// TwinCAT 3 PLC project TestSample
// ProgramVersion: 3.1.4026.28
// libraries:
//   Tc2_Standard, * (Beckhoff Automation GmbH)
//   Tc2_System, * (Beckhoff Automation GmbH)
//   Tc2_TcpIp, * (Beckhoff Automation GmbH)
//   Tc3_Module, * (Beckhoff Automation GmbH)
// project tree:
//   Diagram/ Class Diagram.TcCD (not stored)
//   Generated/DUT_Generated/ ST_VC_InspectionResult.TcDUT, ST_VC_MoveToPositionArgs.TcDUT, ST_VC_MoveToPositionResult.TcDUT, ST_VC_ReportModuleStateArgs.TcDUT
//   Generated/GVLs_Generated/ GVL_VC_Methods.TcGVL
//   Generated/POU_Generated/ VC_Call_StartInspection.TcPOU, VC_Handle_MoveToPosition.TcPOU, VC_Handle_ReportModuleState.TcPOU
//   Library/DUT/ E_VC_LinkState.TcDUT, E_VC_MsgType.TcDUT, E_VC_SlotState.TcDUT, ST_VC_CtrlMsg.TcDUT, ST_VC_Diag.TcDUT, ST_VC_Header.TcDUT, ST_VC_InSlot.TcDUT, ST_VC_LinkData.TcDUT, ST_VC_MethodInfo.TcDUT, ST_VC_OutSlot.TcDUT
//   Library/GVL/ GVL_VC_Param.TcGVL
//   Library/POU/ VC_CancelOutSlot.TcPOU, VC_CompleteInSlot.TcPOU, VC_DecodeHeader.TcPOU, VC_EncodeHeader.TcPOU, VC_Framer.TcPOU, VC_GetBool.TcPOU, VC_GetFloat32.TcPOU, VC_GetFloat32Array.TcPOU, VC_GetFloat64.TcPOU, VC_GetInt16.TcPOU, VC_GetInt32.TcPOU, VC_GetInt64.TcPOU, VC_GetInt8.TcPOU, VC_GetRaw.TcPOU, VC_GetString.TcPOU, VC_GetUInt16.TcPOU, VC_GetUInt32.TcPOU, VC_GetUInt64.TcPOU, VC_GetUInt8.TcPOU, VC_IsCallable.TcPOU, VC_Link.TcPOU, VC_MethodIndex.TcPOU, VC_PutBool.TcPOU, VC_PutFloat32.TcPOU, VC_PutFloat32Array.TcPOU, VC_PutFloat64.TcPOU, VC_PutInt16.TcPOU, VC_PutInt32.TcPOU, VC_PutInt64.TcPOU, VC_PutInt8.TcPOU, VC_PutRaw.TcPOU, VC_PutString.TcPOU, VC_PutUInt16.TcPOU, VC_PutUInt32.TcPOU, VC_PutUInt64.TcPOU, VC_PutUInt8.TcPOU, VC_ReleaseOutSlot.TcPOU, VC_ReserveOutSlot.TcPOU, VC_SubmitOutSlot.TcPOU, VC_TakeInSlot.TcPOU, VC_Transport.TcPOU
//   / PlcTask.TcTTO
//   POUs/ MAIN.TcPOU
//   Test/GVL/ GVL_VC.TcGVL
//   Test/POU/ FB_VC_LinkTest.TcPOU, MAIN_1.TcPOU
// real-time tasks:
//   TASK PlcTask: cycle T#10ms, priority 20, ADS port 350

CONFIGURATION TestSample
    RESOURCE PLC ON TwinCAT3
        TASK PlcTask(INTERVAL := T#10ms, PRIORITY := 20);
    END_RESOURCE
END_CONFIGURATION

// ---- Generated/DUT_Generated/ST_VC_InspectionResult.TcDUT
TYPE ST_VC_InspectionResult :
STRUCT
    Pass          : BOOL;
    ErrorCode     : DINT;
    MeasuredCount : UINT;
    Measured      : ARRAY[0..15] OF REAL;
END_STRUCT
END_TYPE

// ---- Generated/DUT_Generated/ST_VC_MoveToPositionArgs.TcDUT
TYPE ST_VC_MoveToPositionArgs :
STRUCT
    Position : LREAL;
END_STRUCT
END_TYPE

// ---- Generated/DUT_Generated/ST_VC_MoveToPositionResult.TcDUT
TYPE ST_VC_MoveToPositionResult :
STRUCT
    Accepted : BOOL;
END_STRUCT
END_TYPE

// ---- Generated/DUT_Generated/ST_VC_ReportModuleStateArgs.TcDUT
TYPE ST_VC_ReportModuleStateArgs :
STRUCT
    State   : UINT;     // PackML state from VisionCore
    AlarmId : DINT;
END_STRUCT
END_TYPE

// ---- Library/DUT/E_VC_LinkState.TcDUT
TYPE E_VC_LinkState :
(
    VC_LS_DISABLED   := 0,
    VC_LS_CONNECTING := 1,   // PLC connects actively (VisionCore mode Listen)
    VC_LS_LISTENING  := 2,   // PLC waits for connection (VisionCore mode Connect)
    VC_LS_HELLO      := 3,   // Hello sent, waiting for HelloAck
    VC_LS_ONLINE     := 4,
    VC_LS_CLOSING    := 5,
    VC_LS_WAIT_RETRY := 6
) UINT;
END_TYPE

// ---- Library/DUT/E_VC_MsgType.TcDUT
TYPE E_VC_MsgType :
// Deliberately NOT {attribute 'strict'}: values are compared with the USINT header field.
(
    VC_MT_HELLO     := 1,
    VC_MT_HELLO_ACK := 2,
    VC_MT_REQUEST   := 3,
    VC_MT_RESPONSE  := 4,
    VC_MT_CANCEL    := 5,
    VC_MT_HEARTBEAT := 6
) USINT;
END_TYPE

// ---- Library/DUT/E_VC_SlotState.TcDUT
TYPE E_VC_SlotState :
(
    VC_SS_FREE           := 0,
    VC_SS_RESERVED       := 1,   // Out: block owns slot
    VC_SS_TX_PENDING     := 2,   // Out: request ready to send
    VC_SS_SENT           := 3,   // Out: request sent, waiting for response
    VC_SS_CANCEL_PENDING := 4,   // Out: Cancel must be sent
    VC_SS_DONE           := 5,   // Out: response or error available
    VC_SS_REQUEST        := 10,  // In:  request received, no handler yet
    VC_SS_IN_PROGRESS    := 11,  // In:  handler working
    VC_SS_RESPONSE_READY := 12   // In:  response ready to send
) UINT;
END_TYPE

// ---- Library/DUT/ST_VC_CtrlMsg.TcDUT
TYPE ST_VC_CtrlMsg :              // Cancel or error response without payload
STRUCT
    MessageType : E_VC_MsgType;
    MethodId    : UINT;
    CallId      : UDINT;
    Status      : UINT;
END_STRUCT
END_TYPE

// ---- Library/DUT/ST_VC_Diag.TcDUT
TYPE ST_VC_Diag :
STRUCT
    RxMessages          : UDINT;
    TxMessages          : UDINT;
    ProtocolErrors      : UDINT;
    Reconnects          : UDINT;
    CallTimeouts        : UDINT;
    RejectedCalls       : UDINT;
    LastErrorId         : UINT;
    LastErrorMs         : UDINT;
    LastTransportStatus : DWORD;  // raw nErrId of the Tc2_TcpIp block
END_STRUCT
END_TYPE

// ---- Library/DUT/ST_VC_Header.TcDUT
{attribute 'pack_mode' := '1'}
TYPE ST_VC_Header :
STRUCT
    Magic           : UINT;    // 16#5643, little-endian on the wire (43 56)
    ProtocolVersion : USINT;   // 1
    MessageType     : USINT;   // E_VC_MsgType
    Flags           : UINT;    // reserved, 0
    MethodId        : UINT;    // 0 for Hello / Heartbeat
    CallId          : UDINT;   // bit 31 = 1: call from VisionCore
    PayloadLength   : UDINT;
    Status          : UINT;    // response status, else 0
    Reserved        : UINT;
END_STRUCT
END_TYPE

// ---- Library/DUT/ST_VC_InSlot.TcDUT
TYPE ST_VC_InSlot :               // App calls PLC
STRUCT
    State           : E_VC_SlotState;
    MethodIndex     : UINT;
    CallId          : UDINT;
    ReceivedMs      : UDINT;
    CancelRequested : BOOL;
    Status          : UINT;
    PayloadLen      : UDINT;
    Payload         : ARRAY[0..VC_MAX_PAYLOAD - 1] OF BYTE;  // arguments first, then result
END_STRUCT
END_TYPE

// ---- Library/DUT/ST_VC_LinkData.TcDUT
TYPE ST_VC_LinkData :
STRUCT
    // State
    State          : E_VC_LinkState;
    Online         : BOOL;
    NowMs          : UDINT;      // time base, set by VC_Link every cycle
    StateSinceMs   : UDINT;
    LastRxMs       : UDINT;
    LastTxMs       : UDINT;
    NextCallId     : UDINT;      // 1 .. 16#7FFFFFFF, bit 31 always 0

    // Release from HelloAck and handler presence, index = method index
    MethodState    : ARRAY[0..VC_MAX_METHODS - 1] OF USINT;  // 0 unknown, 1 released, 2 hash, 3 not allowed
    HandlerSeenMs  : ARRAY[0..VC_MAX_METHODS - 1] OF UDINT;

    // Call slots
    OutSlots       : ARRAY[0..VC_MAX_CALLS - 1] OF ST_VC_OutSlot;
    InSlots        : ARRAY[0..VC_MAX_CALLS - 1] OF ST_VC_InSlot;
    NextOutSend    : UINT;       // round robin for sending

    // Control messages
    CtrlQueue      : ARRAY[0..VC_CTRL_QUEUE - 1] OF ST_VC_CtrlMsg;
    CtrlHead       : UINT;
    CtrlCount      : UINT;

    // Buffers
    RxBuffer       : ARRAY[0..VC_RX_BUFFER - 1] OF BYTE;
    RxFill         : UDINT;
    TxFrame        : ARRAY[0..VC_HEADER_LEN + VC_MAX_PAYLOAD - 1] OF BYTE;

    // Diagnostics
    Diag           : ST_VC_Diag;
END_STRUCT
END_TYPE

// ---- Library/DUT/ST_VC_MethodInfo.TcDUT
TYPE ST_VC_MethodInfo :
STRUCT
    MethodId  : UINT;
    Hash      : UDINT;   // CRC-32 of canonical signature (generated)
    Provider  : USINT;   // 0 = App, 1 = Plc
    TimeoutMs : UDINT;
    ArgsLen   : UDINT;   // request payload length
    ResultLen : UDINT;   // response payload length at status 0
END_STRUCT
END_TYPE

// ---- Library/DUT/ST_VC_OutSlot.TcDUT
TYPE ST_VC_OutSlot :              // PLC calls App
STRUCT
    State        : E_VC_SlotState;
    MethodIndex  : UINT;
    CallId       : UDINT;
    StartMs      : UDINT;
    TimeoutMs    : UDINT;
    OwnerSeenMs  : UDINT;         // last call of owning VC_Call_* block
    Status       : UINT;
    PayloadLen   : UDINT;
    Payload      : ARRAY[0..VC_MAX_PAYLOAD - 1] OF BYTE;  // arguments first, then result
END_STRUCT
END_TYPE

// ---- Generated/GVLs_Generated/GVL_VC_Methods.TcGVL
VAR_GLOBAL CONSTANT
// ===== GENERATED PART (normally written by vcgen) - hand-written stand-in for testing =====
// Hash = CRC-32 (IEEE, as zlib) over the canonical signature, SPS-Konzept 4.5:
//   10|StartInspection|App|UInt16,String32|Bool,Int32,UInt16,Float32[16]
//   500|ReportModuleState|Plc|UInt16,Int32|
//   600|MoveToPosition|Plc|Float64|Bool
// ASSUMPTION: VisionCore computes the same CRC variant and string. If not, HelloAck returns
// MethodState 2 and calls fail with ErrorId 2 -> copy the hashes from the VisionCore build.
    VC_METHOD_COUNT            : UINT := 3;

    // Method index = position in VC_METHODS (used by all blocks)
    VC_IDX_START_INSPECTION    : UINT := 0;
    VC_IDX_REPORT_MODULE_STATE : UINT := 1;
    VC_IDX_MOVE_TO_POSITION    : UINT := 2;

    // ASSUMPTION: project interface name, confirm with VisionCore configuration
    VC_INTERFACES : ARRAY[0..3] OF STRING(47) := ['VisionCore.Platform', 'Stent.Line1', '', ''];

    VC_METHODS : ARRAY[0..VC_MAX_METHODS - 1] OF ST_VC_MethodInfo := [
        // StartInspection: args UInt16 + String32 = 34; result Bool+Int32+UInt16+16xFloat32 = 71
        (MethodId := 10,  Hash := 16#A1EFD4EB, Provider := 0, TimeoutMs := 10000, ArgsLen := 34, ResultLen := 71),
        // ReportModuleState: args UInt16 + Int32 = 6; no result
        (MethodId := 500, Hash := 16#18245D80, Provider := 1, TimeoutMs := 200,   ArgsLen := 6,  ResultLen := 0),
        // MoveToPosition: args Float64 = 8; result Bool = 1. ASSUMPTION: timeout 5000 ms
        (MethodId := 600, Hash := 16#689DF4EB, Provider := 1, TimeoutMs := 5000,  ArgsLen := 8,  ResultLen := 1)
    ];
END_VAR

// ---- Library/GVL/GVL_VC_Param.TcGVL
VAR_GLOBAL CONSTANT
    // ---- Protocol (fixed, SPS-Konzept section 5) ----
    VC_MAGIC              : UINT  := 16#5643;   // 'VC'
    VC_PROTOCOL_VERSION   : USINT := 1;
    VC_HEADER_LEN         : UDINT := 20;
    VC_HELLO_ACK_LEN      : UDINT := 65;        // Accepted + 64 x MethodState
    VC_PROVIDER_APP       : USINT := 0;
    VC_PROVIDER_PLC       : USINT := 1;

    // ---- Parameters (Bausteindesign section 3) ----
    VC_MAX_PAYLOAD        : UDINT := 4096;
    VC_MAX_CALLS          : UINT  := 8;
    VC_MAX_METHODS        : UINT  := 64;        // must stay 64: Hello/HelloAck carry 64 entries
    VC_RX_BUFFER          : UDINT := 2 * (VC_HEADER_LEN + VC_MAX_PAYLOAD);
    VC_CTRL_QUEUE         : UINT  := 16;
    VC_MSG_PER_CYCLE      : UINT  := 4;
    VC_HELLO_TIMEOUT_MS   : UDINT := 5000;
    VC_HEARTBEAT_MS       : UDINT := 1000;
    VC_WATCHDOG_MS        : UDINT := 3000;
    VC_RETRY_MS           : UDINT := 2000;
    VC_OWNER_TIMEOUT_MS   : UDINT := 1000;

    // ---- Status codes (SPS-Konzept 5.7) ----
    VC_STATUS_OK                  : UINT := 0;
    VC_STATUS_UNKNOWN_METHOD      : UINT := 1;
    VC_STATUS_METHOD_INCOMPATIBLE : UINT := 2;
    VC_STATUS_NOT_ALLOWED         : UINT := 3;
    VC_STATUS_INVALID_PAYLOAD     : UINT := 4;
    VC_STATUS_BUSY                : UINT := 5;
    VC_STATUS_CANCELLED           : UINT := 6;
    VC_STATUS_TIMEOUT             : UINT := 7;
    VC_STATUS_CONNECTION_LOST     : UINT := 8;
    VC_STATUS_INTERNAL_ERROR      : UINT := 9;

    // ---- VC_Link.ErrorId (Bausteindesign section 8) ----
    VC_ERR_CONNECT         : UINT := 1;   // connect / listen / accept failed
    VC_ERR_HELLO_TIMEOUT   : UINT := 2;   // no HelloAck in time
    VC_ERR_HELLO_REJECTED  : UINT := 3;   // HelloAck Accepted = FALSE
    VC_ERR_PROTOCOL        : UINT := 4;   // invalid header / unexpected message
    VC_ERR_WATCHDOG        : UINT := 5;   // nothing received
    VC_ERR_SEND            : UINT := 6;
    VC_ERR_RECEIVE         : UINT := 7;
END_VAR

// ---- Test/GVL/GVL_VC.TcGVL
VAR_GLOBAL
    LinkData : ST_VC_LinkData;   // one per VisionCore connection, ~80 KB
END_VAR

// ---- Library/POU/VC_Link.TcPOU
FUNCTION_BLOCK VC_Link
// Central block: one instance per VisionCore connection, called every cycle,
// BEFORE all VC_Call_* / VC_Handle_* blocks that use the same ST_VC_LinkData (same task).
VAR_INPUT
    Enable        : BOOL;
    Mode          : INT;           // 0 = connect actively, 1 = wait for connection
    RemoteAddress : STRING(15);    // Mode = 0
    RemotePort    : UINT := 5100;  // Mode = 0
    LocalPort     : UINT := 5100;  // Mode = 1
    ClientId      : STRING(31);
END_VAR
VAR_IN_OUT
    Link          : ST_VC_LinkData;
END_VAR
VAR_OUTPUT
    Connected     : BOOL;          // TCP connection up
    Online        : BOOL;          // HelloAck received
    Restricted    : BOOL;          // at least one method not released
    Error         : BOOL;          // stays set until ONLINE again
    ErrorId       : UINT;          // VC_ERR_*
    State         : E_VC_LinkState;
END_VAR
VAR
    fbTransport   : VC_Transport;
    fbFramer      : VC_Framer;
    bSendReq      : BOOL;          // frame in TxFrame, waiting for transport to take it
    nTxLen        : UDINT;
    bHelloSent    : BOOL;
    nIdx          : UINT;
END_VAR

// ---- 1. Time base ----
Link.NowMs := TIME_TO_UDINT(TIME());

// ---- 2./3. Transport: connect, accept, close, send, receive ----
fbTransport(
    Open          := (Link.State = VC_LS_CONNECTING) OR (Link.State = VC_LS_LISTENING)
                     OR (Link.State = VC_LS_HELLO) OR (Link.State = VC_LS_ONLINE),
    Mode          := Mode,
    RemoteAddress := RemoteAddress,
    RemotePort    := RemotePort,
    LocalPort     := LocalPort,
    SendRequest   := bSendReq,
    SendLen       := nTxLen,
    Link          := Link);
IF fbTransport.SendBusy THEN
    bSendReq := FALSE;                 // transport has taken the frame
END_IF
IF fbTransport.Error THEN
    Link.Diag.LastTransportStatus := fbTransport.Status;
END_IF

// ---- Connection state machine ----
CASE Link.State OF
VC_LS_DISABLED:
    IF Enable THEN
        IF Mode = 0 THEN
            THIS^.GotoState(stLink := Link, NewState := VC_LS_CONNECTING);
        ELSE
            THIS^.GotoState(stLink := Link, NewState := VC_LS_LISTENING);
        END_IF
    END_IF

VC_LS_CONNECTING, VC_LS_LISTENING:
    IF NOT Enable THEN
        THIS^.GotoState(stLink := Link, NewState := VC_LS_CLOSING);
    ELSIF fbTransport.Error THEN
        THIS^.SetError(stLink := Link, Id := VC_ERR_CONNECT);
        THIS^.GotoState(stLink := Link, NewState := VC_LS_CLOSING);   // releases handles, then WAIT_RETRY
    ELSIF fbTransport.Connected THEN
        THIS^.GotoState(stLink := Link, NewState := VC_LS_HELLO);
    END_IF

VC_LS_HELLO, VC_LS_ONLINE:
    IF NOT Enable THEN
        THIS^.GotoState(stLink := Link, NewState := VC_LS_CLOSING);
    ELSIF fbTransport.Error THEN
        THIS^.SetError(stLink := Link, Id := fbTransport.ErrorId);
        THIS^.GotoState(stLink := Link, NewState := VC_LS_CLOSING);
    ELSIF NOT fbTransport.Connected THEN
        THIS^.SetError(stLink := Link, Id := VC_ERR_RECEIVE);
        THIS^.GotoState(stLink := Link, NewState := VC_LS_CLOSING);
    END_IF

VC_LS_CLOSING:
    IF fbTransport.Idle THEN
        IF Enable THEN
            THIS^.GotoState(stLink := Link, NewState := VC_LS_WAIT_RETRY);
        ELSE
            THIS^.GotoState(stLink := Link, NewState := VC_LS_DISABLED);
        END_IF
    END_IF

VC_LS_WAIT_RETRY:
    IF NOT Enable THEN
        THIS^.GotoState(stLink := Link, NewState := VC_LS_DISABLED);
    ELSIF (Link.NowMs - Link.StateSinceMs) >= VC_RETRY_MS THEN
        IF Mode = 0 THEN
            THIS^.GotoState(stLink := Link, NewState := VC_LS_CONNECTING);
        ELSE
            THIS^.GotoState(stLink := Link, NewState := VC_LS_LISTENING);
        END_IF
    END_IF
END_CASE

// ---- 4. Process messages ----
IF (Link.State = VC_LS_HELLO) OR (Link.State = VC_LS_ONLINE) THEN
    THIS^.ProcessMessages(stLink := Link);
END_IF

// ---- 5. Deadlines ----
IF (Link.State = VC_LS_HELLO) OR (Link.State = VC_LS_ONLINE) THEN
    THIS^.CheckDeadlines(stLink := Link);
END_IF

// ---- 6. Schedule at most one message ----
IF (Link.State = VC_LS_HELLO) OR (Link.State = VC_LS_ONLINE) THEN
    THIS^.ScheduleSend(stLink := Link);
END_IF

// ---- 7. Outputs ----
Connected  := fbTransport.Connected;
Online     := Link.Online;
State      := Link.State;
Restricted := FALSE;
IF Link.Online THEN
    nIdx := 0;
    WHILE (nIdx < VC_METHOD_COUNT) AND (nIdx < VC_MAX_METHODS) DO
        IF Link.MethodState[nIdx] <> 1 THEN
            Restricted := TRUE;
        END_IF
        nIdx := nIdx + 1;
    END_WHILE
END_IF

METHOD PRIVATE BuildHello : UDINT
// Bausteindesign 7.3: 32 + 4 x 48 + 2 + 64 x 6 = 610 bytes payload
VAR_IN_OUT
    stLink : ST_VC_LinkData;
END_VAR
VAR
    nPos : UDINT;
    k    : UINT;
END_VAR
nPos := VC_HEADER_LEN;
VC_PutString(Buf := stLink.TxFrame, Pos := nPos, Value := ClientId, Len := 32);
FOR k := 0 TO 3 DO
    VC_PutString(Buf := stLink.TxFrame, Pos := nPos, Value := VC_INTERFACES[k], Len := 48);
END_FOR
VC_PutUInt16(Buf := stLink.TxFrame, Pos := nPos, Value := VC_METHOD_COUNT);
FOR k := 0 TO VC_MAX_METHODS - 1 DO
    VC_PutUInt16(Buf := stLink.TxFrame, Pos := nPos, Value := VC_METHODS[k].MethodId);
    VC_PutUInt32(Buf := stLink.TxFrame, Pos := nPos, Value := VC_METHODS[k].Hash);
END_FOR
BuildHello := nPos - VC_HEADER_LEN;
END_METHOD

METHOD PRIVATE CheckDeadlines
VAR_IN_OUT
    stLink : ST_VC_LinkData;
END_VAR
VAR
    k    : UINT;
    nIdx : UINT;
END_VAR
// Hello timeout / watchdog
IF stLink.State = VC_LS_HELLO THEN
    IF (stLink.NowMs - stLink.StateSinceMs) > VC_HELLO_TIMEOUT_MS THEN
        THIS^.SetError(stLink := stLink, Id := VC_ERR_HELLO_TIMEOUT);
        THIS^.GotoState(stLink := stLink, NewState := VC_LS_CLOSING);
        RETURN;
    END_IF
ELSIF stLink.State = VC_LS_ONLINE THEN
    IF (stLink.NowMs - stLink.LastRxMs) > VC_WATCHDOG_MS THEN
        THIS^.SetError(stLink := stLink, Id := VC_ERR_WATCHDOG);
        THIS^.GotoState(stLink := stLink, NewState := VC_LS_CLOSING);
        RETURN;
    END_IF
END_IF

FOR k := 0 TO VC_MAX_CALLS - 1 DO
    // Out slots: call timeout and orphaned slots
    CASE stLink.OutSlots[k].State OF
    VC_SS_SENT:
        IF (stLink.NowMs - stLink.OutSlots[k].StartMs) > stLink.OutSlots[k].TimeoutMs THEN
            stLink.OutSlots[k].Status := VC_STATUS_TIMEOUT;
            stLink.OutSlots[k].State  := VC_SS_CANCEL_PENDING;
            stLink.Diag.CallTimeouts  := stLink.Diag.CallTimeouts + 1;
        END_IF
    VC_SS_RESERVED, VC_SS_DONE:
        IF (stLink.NowMs - stLink.OutSlots[k].OwnerSeenMs) > VC_OWNER_TIMEOUT_MS THEN
            stLink.OutSlots[k].State      := VC_SS_FREE;
            stLink.OutSlots[k].Status     := VC_STATUS_OK;
            stLink.OutSlots[k].PayloadLen := 0;
        END_IF
    END_CASE

    // In slots: released without answer after 2 x method timeout
    CASE stLink.InSlots[k].State OF
    VC_SS_REQUEST, VC_SS_IN_PROGRESS:
        nIdx := stLink.InSlots[k].MethodIndex;
        IF (stLink.NowMs - stLink.InSlots[k].ReceivedMs) > (2 * VC_METHODS[nIdx].TimeoutMs) THEN
            stLink.InSlots[k].State           := VC_SS_FREE;
            stLink.InSlots[k].CancelRequested := FALSE;
        END_IF
    END_CASE
END_FOR
END_METHOD

METHOD PRIVATE EnqueueCtrl : BOOL
VAR_IN_OUT
    stLink   : ST_VC_LinkData;
END_VAR
VAR_INPUT
    MsgType  : E_VC_MsgType;
    MethodId : UINT;
    CallId   : UDINT;
    Status   : UINT;
END_VAR
VAR
    nTail : UINT;
END_VAR
IF stLink.CtrlCount >= VC_CTRL_QUEUE THEN
    EnqueueCtrl := FALSE;                                  // queue full: VisionCore runs into its timeout
    RETURN;
END_IF
nTail := (stLink.CtrlHead + stLink.CtrlCount) MOD VC_CTRL_QUEUE;
stLink.CtrlQueue[nTail].MessageType := MsgType;
stLink.CtrlQueue[nTail].MethodId    := MethodId;
stLink.CtrlQueue[nTail].CallId      := CallId;
stLink.CtrlQueue[nTail].Status      := Status;
stLink.CtrlCount := stLink.CtrlCount + 1;
EnqueueCtrl := TRUE;
END_METHOD

METHOD PRIVATE GotoState
VAR_IN_OUT
    stLink   : ST_VC_LinkData;
END_VAR
VAR_INPUT
    NewState : E_VC_LinkState;
END_VAR
stLink.State        := NewState;
stLink.StateSinceMs := stLink.NowMs;

CASE NewState OF
VC_LS_HELLO:
    stLink.RxFill := 0;
    bHelloSent    := FALSE;
VC_LS_ONLINE:
    stLink.Online   := TRUE;
    stLink.LastRxMs := stLink.NowMs;
    Error           := FALSE;
    ErrorId         := 0;
VC_LS_CLOSING:
    THIS^.HandleConnectionLoss(stLink := stLink);
VC_LS_WAIT_RETRY:
    stLink.Diag.Reconnects := stLink.Diag.Reconnects + 1;
END_CASE
END_METHOD

METHOD PRIVATE HandleCancel
// Cancel from VisionCore. Not yet taken by a handler -> answer Cancelled directly.
VAR_IN_OUT
    stLink : ST_VC_LinkData;
END_VAR
VAR_INPUT
    Hdr    : ST_VC_Header;
END_VAR
VAR
    k : UINT;
END_VAR
FOR k := 0 TO VC_MAX_CALLS - 1 DO
    IF stLink.InSlots[k].CallId = Hdr.CallId THEN
        CASE stLink.InSlots[k].State OF
        VC_SS_REQUEST:
            stLink.InSlots[k].Status     := VC_STATUS_CANCELLED;
            stLink.InSlots[k].PayloadLen := 0;
            stLink.InSlots[k].State      := VC_SS_RESPONSE_READY;
            RETURN;
        VC_SS_IN_PROGRESS:
            stLink.InSlots[k].CancelRequested := TRUE;   // handler answers Cancelled or regular
            RETURN;
        END_CASE
    END_IF
END_FOR
END_METHOD

METHOD PRIVATE HandleConnectionLoss
// Bausteindesign section 5: "Verbindungsabbruch behandeln" (handle connection loss)
VAR_IN_OUT
    stLink : ST_VC_LinkData;
END_VAR
VAR
    k : UINT;
END_VAR
stLink.Online := FALSE;
FOR k := 0 TO VC_MAX_METHODS - 1 DO
    stLink.MethodState[k] := 0;
END_FOR
FOR k := 0 TO VC_MAX_CALLS - 1 DO
    CASE stLink.OutSlots[k].State OF
    VC_SS_TX_PENDING, VC_SS_SENT, VC_SS_CANCEL_PENDING:
        stLink.OutSlots[k].Status     := VC_STATUS_CONNECTION_LOST;
        stLink.OutSlots[k].PayloadLen := 0;
        stLink.OutSlots[k].State      := VC_SS_DONE;
    END_CASE
    stLink.InSlots[k].State           := VC_SS_FREE;   // VisionCore reports the loss itself
    stLink.InSlots[k].CancelRequested := FALSE;
END_FOR
stLink.CtrlHead  := 0;
stLink.CtrlCount := 0;
stLink.RxFill    := 0;
bSendReq         := FALSE;
END_METHOD

METHOD PRIVATE HandleHelloAck
VAR_IN_OUT
    stLink : ST_VC_LinkData;
END_VAR
VAR_INPUT
    Hdr    : ST_VC_Header;
END_VAR
VAR
    k : UINT;
END_VAR
// Only valid in HELLO and with exactly 65 bytes payload
IF (stLink.State <> VC_LS_HELLO) OR (Hdr.PayloadLength <> VC_HELLO_ACK_LEN) THEN
    THIS^.SetError(stLink := stLink, Id := VC_ERR_PROTOCOL);
    THIS^.GotoState(stLink := stLink, NewState := VC_LS_CLOSING);
    RETURN;
END_IF

IF stLink.RxBuffer[VC_HEADER_LEN] = 0 THEN                 // Accepted = FALSE
    THIS^.SetError(stLink := stLink, Id := VC_ERR_HELLO_REJECTED);
    THIS^.GotoState(stLink := stLink, NewState := VC_LS_CLOSING);
    RETURN;
END_IF

FOR k := 0 TO VC_MAX_METHODS - 1 DO
    stLink.MethodState[k] := BYTE_TO_USINT(stLink.RxBuffer[VC_HEADER_LEN + 1 + k]);
END_FOR
THIS^.GotoState(stLink := stLink, NewState := VC_LS_ONLINE);
END_METHOD

METHOD PRIVATE HandleRequest
// Request from VisionCore: checks from Bausteindesign 6.2, then occupy an in slot.
VAR_IN_OUT
    stLink : ST_VC_LinkData;
END_VAR
VAR_INPUT
    Hdr    : ST_VC_Header;
END_VAR
VAR
    k       : UINT;
    nIdx    : INT;
    nSlot   : INT;
    nStatus : UINT;
END_VAR
nSlot   := -1;
nStatus := VC_STATUS_OK;
nIdx    := VC_MethodIndex(MethodId := Hdr.MethodId, Provider := VC_PROVIDER_PLC);

IF nIdx < 0 THEN
    nStatus := VC_STATUS_UNKNOWN_METHOD;
ELSIF stLink.MethodState[nIdx] <> 1 THEN
    nStatus := VC_STATUS_METHOD_INCOMPATIBLE;
ELSIF (stLink.NowMs - stLink.HandlerSeenMs[nIdx]) >= VC_OWNER_TIMEOUT_MS THEN
    nStatus := VC_STATUS_UNKNOWN_METHOD;                   // no active VC_Handle_* instance
ELSIF Hdr.PayloadLength <> VC_METHODS[nIdx].ArgsLen THEN
    nStatus := VC_STATUS_INVALID_PAYLOAD;
ELSE
    FOR k := 0 TO VC_MAX_CALLS - 1 DO
        IF stLink.InSlots[k].State = VC_SS_FREE THEN
            nSlot := UINT_TO_INT(k);
            EXIT;
        END_IF
    END_FOR
    IF nSlot < 0 THEN
        nStatus := VC_STATUS_BUSY;
    END_IF
END_IF

IF nStatus <> VC_STATUS_OK THEN
    THIS^.EnqueueCtrl(stLink := stLink, MsgType := VC_MT_RESPONSE,
                      MethodId := Hdr.MethodId, CallId := Hdr.CallId, Status := nStatus);
    stLink.Diag.RejectedCalls := stLink.Diag.RejectedCalls + 1;
    RETURN;
END_IF

stLink.InSlots[nSlot].MethodIndex     := INT_TO_UINT(nIdx);
stLink.InSlots[nSlot].CallId          := Hdr.CallId;
stLink.InSlots[nSlot].ReceivedMs      := stLink.NowMs;
stLink.InSlots[nSlot].CancelRequested := FALSE;
stLink.InSlots[nSlot].Status          := VC_STATUS_OK;
stLink.InSlots[nSlot].PayloadLen      := Hdr.PayloadLength;
IF Hdr.PayloadLength > 0 THEN
    MEMCPY(destAddr := ADR(stLink.InSlots[nSlot].Payload),
           srcAddr  := ADR(stLink.RxBuffer[VC_HEADER_LEN]),
           n        := Hdr.PayloadLength);
END_IF
stLink.InSlots[nSlot].State := VC_SS_REQUEST;
END_METHOD

METHOD PRIVATE HandleResponse
// Response to a PLC call: match out slot in SENT by CallId; late responses are discarded.
VAR_IN_OUT
    stLink : ST_VC_LinkData;
END_VAR
VAR_INPUT
    Hdr    : ST_VC_Header;
END_VAR
VAR
    k     : UINT;
    nSlot : INT;
    nIdx  : UINT;
END_VAR
nSlot := -1;
FOR k := 0 TO VC_MAX_CALLS - 1 DO
    IF (stLink.OutSlots[k].State = VC_SS_SENT) AND (stLink.OutSlots[k].CallId = Hdr.CallId) THEN
        nSlot := UINT_TO_INT(k);
        EXIT;
    END_IF
END_FOR
IF nSlot < 0 THEN
    RETURN;                                                // cancelled / timed out / unknown -> drop
END_IF

nIdx := stLink.OutSlots[nSlot].MethodIndex;
IF Hdr.Status = VC_STATUS_OK THEN
    IF (Hdr.MethodId = VC_METHODS[nIdx].MethodId) AND (Hdr.PayloadLength = VC_METHODS[nIdx].ResultLen) THEN
        IF Hdr.PayloadLength > 0 THEN
            MEMCPY(destAddr := ADR(stLink.OutSlots[nSlot].Payload),
                   srcAddr  := ADR(stLink.RxBuffer[VC_HEADER_LEN]),
                   n        := Hdr.PayloadLength);
        END_IF
        stLink.OutSlots[nSlot].PayloadLen := Hdr.PayloadLength;
        stLink.OutSlots[nSlot].Status     := VC_STATUS_OK;
    ELSE
        stLink.OutSlots[nSlot].PayloadLen := 0;
        stLink.OutSlots[nSlot].Status     := VC_STATUS_INVALID_PAYLOAD;
    END_IF
ELSE
    stLink.OutSlots[nSlot].PayloadLen := 0;
    stLink.OutSlots[nSlot].Status     := Hdr.Status;
END_IF
stLink.OutSlots[nSlot].State := VC_SS_DONE;
END_METHOD

METHOD PRIVATE ProcessMessages
// Bausteindesign 7.1: at most VC_MSG_PER_CYCLE messages per cycle
VAR_IN_OUT
    stLink : ST_VC_LinkData;
END_VAR
VAR
    k     : UINT;
    stHdr : ST_VC_Header;
END_VAR
FOR k := 1 TO VC_MSG_PER_CYCLE DO
    fbFramer(Link := stLink);
    IF NOT fbFramer.MessageAvailable THEN
        EXIT;
    END_IF
    IF fbFramer.ProtocolError THEN
        THIS^.SetError(stLink := stLink, Id := VC_ERR_PROTOCOL);
        THIS^.GotoState(stLink := stLink, NewState := VC_LS_CLOSING);
        EXIT;
    END_IF

    stHdr := fbFramer.Header;
    stLink.LastRxMs := stLink.NowMs;                       // resets the watchdog
    stLink.Diag.RxMessages := stLink.Diag.RxMessages + 1;

    CASE stHdr.MessageType OF
    VC_MT_HELLO_ACK:
        THIS^.HandleHelloAck(stLink := stLink, Hdr := stHdr);
    VC_MT_HEARTBEAT:
        ;                                                  // watchdog already reset
    VC_MT_RESPONSE:
        THIS^.HandleResponse(stLink := stLink, Hdr := stHdr);
    VC_MT_REQUEST:
        THIS^.HandleRequest(stLink := stLink, Hdr := stHdr);
    VC_MT_CANCEL:
        THIS^.HandleCancel(stLink := stLink, Hdr := stHdr);
    ELSE                                                   // Hello from App is not allowed
        THIS^.SetError(stLink := stLink, Id := VC_ERR_PROTOCOL);
        THIS^.GotoState(stLink := stLink, NewState := VC_LS_CLOSING);
    END_CASE

    IF stLink.State = VC_LS_CLOSING THEN
        EXIT;                                              // buffer is cleared by HandleConnectionLoss
    END_IF
    fbFramer.Consume(stLink := stLink);
END_FOR
END_METHOD

METHOD PRIVATE ScheduleSend
// Bausteindesign 7.2: build exactly one frame by priority when the transport is free.
VAR_IN_OUT
    stLink : ST_VC_LinkData;
END_VAR
VAR
    k     : UINT;
    nSlot : UINT;
    nIdx  : UINT;
    nLen  : UDINT;
    stMsg : ST_VC_CtrlMsg;
END_VAR
IF bSendReq OR fbTransport.SendBusy OR NOT fbTransport.Connected THEN
    RETURN;                                                // TxFrame still in use
END_IF

// 1. Hello
IF stLink.State = VC_LS_HELLO THEN
    IF NOT bHelloSent THEN
        nLen := THIS^.BuildHello(stLink := stLink);
        THIS^.StartFrame(stLink := stLink, MsgType := VC_MT_HELLO, MethodId := 0, CallId := 0,
                         Status := VC_STATUS_OK, PayloadLen := nLen);
        bHelloSent := TRUE;
    END_IF
    RETURN;
END_IF
IF stLink.State <> VC_LS_ONLINE THEN
    RETURN;
END_IF

// 2. Control messages (error responses)
IF stLink.CtrlCount > 0 THEN
    stMsg := stLink.CtrlQueue[stLink.CtrlHead];
    stLink.CtrlHead  := (stLink.CtrlHead + 1) MOD VC_CTRL_QUEUE;
    stLink.CtrlCount := stLink.CtrlCount - 1;
    THIS^.StartFrame(stLink := stLink, MsgType := stMsg.MessageType, MethodId := stMsg.MethodId,
                     CallId := stMsg.CallId, Status := stMsg.Status, PayloadLen := 0);
    RETURN;
END_IF

// 3. Out slots CANCEL_PENDING -> Cancel, slot DONE
FOR k := 0 TO VC_MAX_CALLS - 1 DO
    IF stLink.OutSlots[k].State = VC_SS_CANCEL_PENDING THEN
        nIdx := stLink.OutSlots[k].MethodIndex;
        THIS^.StartFrame(stLink := stLink, MsgType := VC_MT_CANCEL, MethodId := VC_METHODS[nIdx].MethodId,
                         CallId := stLink.OutSlots[k].CallId, Status := VC_STATUS_OK, PayloadLen := 0);
        stLink.OutSlots[k].State := VC_SS_DONE;
        RETURN;
    END_IF
END_FOR

// 4. In slots RESPONSE_READY -> Response, slot FREE
FOR k := 0 TO VC_MAX_CALLS - 1 DO
    IF stLink.InSlots[k].State = VC_SS_RESPONSE_READY THEN
        nIdx := stLink.InSlots[k].MethodIndex;
        nLen := 0;
        IF stLink.InSlots[k].Status = VC_STATUS_OK THEN
            nLen := stLink.InSlots[k].PayloadLen;
        END_IF
        IF nLen > 0 THEN
            MEMCPY(destAddr := ADR(stLink.TxFrame[VC_HEADER_LEN]),
                   srcAddr  := ADR(stLink.InSlots[k].Payload), n := nLen);
        END_IF
        THIS^.StartFrame(stLink := stLink, MsgType := VC_MT_RESPONSE, MethodId := VC_METHODS[nIdx].MethodId,
                         CallId := stLink.InSlots[k].CallId, Status := stLink.InSlots[k].Status,
                         PayloadLen := nLen);
        stLink.InSlots[k].State           := VC_SS_FREE;
        stLink.InSlots[k].CancelRequested := FALSE;
        RETURN;
    END_IF
END_FOR

// 5. Out slots TX_PENDING -> Request, round robin from NextOutSend
FOR k := 0 TO VC_MAX_CALLS - 1 DO
    nSlot := (stLink.NextOutSend + k) MOD VC_MAX_CALLS;
    IF stLink.OutSlots[nSlot].State = VC_SS_TX_PENDING THEN
        nIdx := stLink.OutSlots[nSlot].MethodIndex;
        nLen := stLink.OutSlots[nSlot].PayloadLen;
        IF nLen > 0 THEN
            MEMCPY(destAddr := ADR(stLink.TxFrame[VC_HEADER_LEN]),
                   srcAddr  := ADR(stLink.OutSlots[nSlot].Payload), n := nLen);
        END_IF
        THIS^.StartFrame(stLink := stLink, MsgType := VC_MT_REQUEST, MethodId := VC_METHODS[nIdx].MethodId,
                         CallId := stLink.OutSlots[nSlot].CallId, Status := VC_STATUS_OK, PayloadLen := nLen);
        stLink.OutSlots[nSlot].State   := VC_SS_SENT;
        stLink.OutSlots[nSlot].StartMs := stLink.NowMs;
        stLink.NextOutSend := (nSlot + 1) MOD VC_MAX_CALLS;
        RETURN;
    END_IF
END_FOR

// 6. Heartbeat
IF (stLink.NowMs - stLink.LastTxMs) >= VC_HEARTBEAT_MS THEN
    THIS^.StartFrame(stLink := stLink, MsgType := VC_MT_HEARTBEAT, MethodId := 0, CallId := 0,
                     Status := VC_STATUS_OK, PayloadLen := 0);
END_IF
END_METHOD

METHOD PRIVATE SetError
VAR_IN_OUT
    stLink : ST_VC_LinkData;
END_VAR
VAR_INPUT
    Id     : UINT;
END_VAR
Error   := TRUE;
ErrorId := Id;
stLink.Diag.LastErrorId := Id;
stLink.Diag.LastErrorMs := stLink.NowMs;
IF Id = VC_ERR_PROTOCOL THEN
    stLink.Diag.ProtocolErrors := stLink.Diag.ProtocolErrors + 1;
END_IF
END_METHOD

METHOD PRIVATE StartFrame
// Writes the header to TxFrame[0..19] (payload must already be at TxFrame[20..]) and requests sending.
VAR_IN_OUT
    stLink     : ST_VC_LinkData;
END_VAR
VAR_INPUT
    MsgType    : E_VC_MsgType;
    MethodId   : UINT;
    CallId     : UDINT;
    Status     : UINT;
    PayloadLen : UDINT;
END_VAR
VAR
    stHdr : ST_VC_Header;
END_VAR
stHdr.Magic           := VC_MAGIC;
stHdr.ProtocolVersion := VC_PROTOCOL_VERSION;
stHdr.MessageType     := TO_USINT(MsgType);
stHdr.Flags           := 0;
stHdr.MethodId        := MethodId;
stHdr.CallId          := CallId;
stHdr.PayloadLength   := PayloadLen;
stHdr.Status          := Status;
stHdr.Reserved        := 0;
VC_EncodeHeader(Buf := stLink.TxFrame, Hdr := stHdr);

nTxLen   := VC_HEADER_LEN + PayloadLen;
bSendReq := TRUE;
stLink.LastTxMs := stLink.NowMs;
stLink.Diag.TxMessages := stLink.Diag.TxMessages + 1;
END_METHOD

END_FUNCTION_BLOCK

// ---- Library/POU/VC_Transport.TcPOU
FUNCTION_BLOCK VC_Transport
// Platform layer (Beckhoff TF6310 / Tc2_TcpIp). The only block that touches sockets.
// Receive goes via an internal buffer and is appended to Link.RxBuffer when complete,
// so VC_Framer may shift RxBuffer while a receive is in flight.
VAR_INPUT
    Open          : BOOL;          // connect / accept while TRUE, close when FALSE
    Mode          : INT;           // 0 = connect actively, 1 = listen
    RemoteAddress : STRING(15);
    RemotePort    : UINT;
    LocalPort     : UINT;
    SendRequest   : BOOL;          // rising edge: send SendLen bytes of Link.TxFrame
    SendLen       : UDINT;
END_VAR
VAR_IN_OUT
    Link          : ST_VC_LinkData;
END_VAR
VAR_OUTPUT
    Connected     : BOOL;
    SendBusy      : BOOL;
    SendDone      : BOOL;          // one cycle
    ReceivedBytes : UDINT;         // bytes appended this cycle
    Error         : BOOL;          // latched until next rising edge of Open
    ErrorId       : UINT;          // VC_ERR_CONNECT / VC_ERR_SEND / VC_ERR_RECEIVE
    Status        : DWORD;         // raw nErrId
    Idle          : BOOL;          // all handles closed, nothing pending
END_VAR
VAR
    fbConnect     : FB_SocketConnect;
    fbListen      : FB_SocketListen;
    fbAccept      : FB_SocketAccept;
    fbClose       : FB_SocketClose;
    fbSend        : FB_SocketSend;
    fbReceive     : FB_SocketReceive;
    rOpen         : R_TRIG;
    rSend         : R_TRIG;
    hSocket       : T_HSOCKET;
    hListener     : T_HSOCKET;
    bSocketOpen   : BOOL;
    bListenerOpen : BOOL;
    bRecvBusy     : BOOL;
    nStep         : INT;
    aRxTemp       : ARRAY[0..VC_HEADER_LEN + VC_MAX_PAYLOAD - 1] OF BYTE;
END_VAR
VAR CONSTANT
    STEP_IDLE           : INT := 0;
    STEP_CONNECT        : INT := 10;
    STEP_LISTEN         : INT := 20;
    STEP_ACCEPT         : INT := 21;
    STEP_CONNECTED      : INT := 30;
    STEP_CLOSE_SOCKET   : INT := 40;
    STEP_CLOSE_LISTENER : INT := 41;
    STEP_WAIT_PENDING   : INT := 42;
    RX_TEMP_LEN         : UDINT := VC_HEADER_LEN + VC_MAX_PAYLOAD;
    TMO                 : TIME := T#5S;
END_VAR

rOpen(CLK := Open);
rSend(CLK := SendRequest);
SendDone      := FALSE;
ReceivedBytes := 0;

IF rOpen.Q THEN
    Error   := FALSE;
    ErrorId := 0;
    Status  := 0;
END_IF

CASE nStep OF
STEP_IDLE:
    IF Open AND NOT Error THEN
        IF Mode = 0 THEN
            nStep := STEP_CONNECT;
        ELSE
            nStep := STEP_LISTEN;
        END_IF
    END_IF

STEP_CONNECT:
    fbConnect(sSrvNetId := '', sRemoteHost := RemoteAddress, nRemotePort := RemotePort,
              bExecute := TRUE, tTimeout := TMO);
    IF NOT fbConnect.bBusy THEN
        fbConnect(bExecute := FALSE);
        IF fbConnect.bError THEN
            THIS^.RaiseError(Id := VC_ERR_CONNECT, Raw := fbConnect.nErrId);
            nStep := STEP_CLOSE_SOCKET;
        ELSE
            hSocket     := fbConnect.hSocket;
            bSocketOpen := TRUE;
            nStep       := STEP_CONNECTED;
        END_IF
    END_IF

STEP_LISTEN:
    fbListen(sSrvNetId := '', sLocalHost := '', nLocalPort := LocalPort,
             bExecute := TRUE, tTimeout := TMO);
    IF NOT fbListen.bBusy THEN
        fbListen(bExecute := FALSE);
        IF fbListen.bError THEN
            THIS^.RaiseError(Id := VC_ERR_CONNECT, Raw := fbListen.nErrId);
            nStep := STEP_CLOSE_SOCKET;
        ELSE
            hListener     := fbListen.hListener;
            bListenerOpen := TRUE;
            nStep         := STEP_ACCEPT;
        END_IF
    END_IF

STEP_ACCEPT:
    IF NOT Open THEN
        nStep := STEP_CLOSE_SOCKET;
    ELSE
        // Re-triggered every second cycle until a client connects
        fbAccept(sSrvNetId := '', hListener := hListener, bExecute := TRUE, tTimeout := TMO);
        IF NOT fbAccept.bBusy THEN
            fbAccept(bExecute := FALSE);
            IF fbAccept.bError THEN
                THIS^.RaiseError(Id := VC_ERR_CONNECT, Raw := fbAccept.nErrId);
                nStep := STEP_CLOSE_SOCKET;
            ELSIF fbAccept.bAccepted THEN
                hSocket     := fbAccept.hSocket;
                bSocketOpen := TRUE;
                nStep       := STEP_CONNECTED;
            END_IF
        END_IF
    END_IF

STEP_CONNECTED:
    IF NOT Open THEN
        nStep := STEP_CLOSE_SOCKET;
    ELSE
        THIS^.ServiceSend(stLink := Link);
        IF nStep = STEP_CONNECTED THEN
            THIS^.ServiceReceive(stLink := Link);
        END_IF
    END_IF

STEP_CLOSE_SOCKET:
    THIS^.DrainPending();
    IF bSocketOpen THEN
        fbClose(sSrvNetId := '', hSocket := hSocket, bExecute := TRUE, tTimeout := TMO);
        IF NOT fbClose.bBusy THEN
            fbClose(bExecute := FALSE);
            bSocketOpen := FALSE;            // handle is gone even if close reported an error
            nStep := STEP_CLOSE_LISTENER;
        END_IF
    ELSE
        nStep := STEP_CLOSE_LISTENER;
    END_IF

STEP_CLOSE_LISTENER:
    THIS^.DrainPending();
    IF bListenerOpen THEN
        fbClose(sSrvNetId := '', hSocket := hListener, bExecute := TRUE, tTimeout := TMO);
        IF NOT fbClose.bBusy THEN
            fbClose(bExecute := FALSE);
            bListenerOpen := FALSE;
            nStep := STEP_WAIT_PENDING;
        END_IF
    ELSE
        nStep := STEP_WAIT_PENDING;
    END_IF

STEP_WAIT_PENDING:
    THIS^.DrainPending();
    IF NOT (fbSend.bBusy OR fbReceive.bBusy OR fbAccept.bBusy OR fbConnect.bBusy OR fbListen.bBusy) THEN
        SendBusy  := FALSE;
        bRecvBusy := FALSE;
        nStep     := STEP_IDLE;
    END_IF
END_CASE

Connected := (nStep = STEP_CONNECTED);
Idle      := (nStep = STEP_IDLE);

METHOD PRIVATE DrainPending
// Keeps running ADS requests alive with bExecute = FALSE until they finish.
IF fbSend.bBusy THEN fbSend(bExecute := FALSE); END_IF
IF fbReceive.bBusy THEN fbReceive(bExecute := FALSE); END_IF
IF fbAccept.bBusy THEN fbAccept(bExecute := FALSE); END_IF
IF fbConnect.bBusy THEN fbConnect(bExecute := FALSE); END_IF
IF fbListen.bBusy THEN fbListen(bExecute := FALSE); END_IF
END_METHOD

METHOD PRIVATE RaiseError
VAR_INPUT
    Id  : UINT;
    Raw : UDINT;
END_VAR
Error   := TRUE;
ErrorId := Id;
Status  := UDINT_TO_DWORD(Raw);
END_METHOD

METHOD PRIVATE ServiceReceive
VAR_IN_OUT
    stLink : ST_VC_LinkData;
END_VAR
VAR
    nFree : UDINT;
    nRec  : UDINT;
END_VAR
// 1. Poll a running receive
IF bRecvBusy THEN
    fbReceive(bExecute := TRUE);
    IF NOT fbReceive.bBusy THEN
        fbReceive(bExecute := FALSE);
        bRecvBusy := FALSE;
        IF fbReceive.bError THEN
            THIS^.RaiseError(Id := VC_ERR_RECEIVE, Raw := fbReceive.nErrId);
            nStep := STEP_CLOSE_SOCKET;
            RETURN;
        END_IF
        nRec := fbReceive.nRecBytes;
        IF nRec > 0 THEN
            IF (stLink.RxFill + nRec) <= VC_RX_BUFFER THEN
                MEMCPY(destAddr := ADR(stLink.RxBuffer[stLink.RxFill]), srcAddr := ADR(aRxTemp), n := nRec);
                stLink.RxFill := stLink.RxFill + nRec;
                ReceivedBytes := nRec;
            ELSE
                THIS^.RaiseError(Id := VC_ERR_RECEIVE, Raw := 0);   // overflow, cannot happen with valid framing
                nStep := STEP_CLOSE_SOCKET;
                RETURN;
            END_IF
        END_IF
    END_IF
END_IF

// 2. Start the next receive (non-blocking, returns 0 bytes if nothing is there)
IF NOT bRecvBusy THEN
    nFree := MIN(VC_RX_BUFFER - stLink.RxFill, RX_TEMP_LEN);
    IF nFree > 0 THEN
        fbReceive(sSrvNetId := '', hSocket := hSocket, cbLen := nFree,
                  pDest := ADR(aRxTemp), bExecute := TRUE, tTimeout := TMO);
        bRecvBusy := TRUE;
    END_IF
END_IF
END_METHOD

METHOD PRIVATE ServiceSend
VAR_IN_OUT
    stLink : ST_VC_LinkData;
END_VAR
IF SendBusy THEN
    fbSend(bExecute := TRUE);
    IF NOT fbSend.bBusy THEN
        fbSend(bExecute := FALSE);
        SendBusy := FALSE;
        IF fbSend.bError THEN
            THIS^.RaiseError(Id := VC_ERR_SEND, Raw := fbSend.nErrId);
            nStep := STEP_CLOSE_SOCKET;
        ELSE
            SendDone := TRUE;
        END_IF
    END_IF
ELSIF rSend.Q THEN
    IF (SendLen > 0) AND (SendLen <= (VC_HEADER_LEN + VC_MAX_PAYLOAD)) THEN
        fbSend(sSrvNetId := '', hSocket := hSocket, cbLen := SendLen,
               pSrc := ADR(stLink.TxFrame), bExecute := TRUE, tTimeout := TMO);
        SendBusy := TRUE;
    END_IF
END_IF
END_METHOD

END_FUNCTION_BLOCK

// ---- Library/POU/VC_Framer.TcPOU
FUNCTION_BLOCK VC_Framer
// Assembles complete messages from the linear RxBuffer and validates the header.
VAR_IN_OUT
    Link             : ST_VC_LinkData;
END_VAR
VAR_OUTPUT
    MessageAvailable : BOOL;     // complete message at RxBuffer[0], or ProtocolError
    ProtocolError    : BOOL;     // wrong Magic / version / type / length
    Header           : ST_VC_Header;
    MessageLen       : UDINT;    // 20 + PayloadLength
END_VAR

MessageAvailable := FALSE;
ProtocolError    := FALSE;
MessageLen       := 0;

IF Link.RxFill < VC_HEADER_LEN THEN
    RETURN;
END_IF

Header := VC_DecodeHeader(Buf := Link.RxBuffer);

IF (Header.Magic <> VC_MAGIC)
    OR (Header.ProtocolVersion <> VC_PROTOCOL_VERSION)
    OR (Header.MessageType < 1) OR (Header.MessageType > 6)
    OR (Header.PayloadLength > VC_MAX_PAYLOAD)
THEN
    ProtocolError    := TRUE;
    MessageAvailable := TRUE;
    RETURN;
END_IF

MessageLen       := VC_HEADER_LEN + Header.PayloadLength;
MessageAvailable := (Link.RxFill >= MessageLen);

METHOD PUBLIC Consume : BOOL
// Removes the current message from RxBuffer and shifts the remaining bytes to index 0.
VAR_IN_OUT
    stLink : ST_VC_LinkData;
END_VAR
Consume := FALSE;
IF (MessageLen = 0) OR (MessageLen > stLink.RxFill) THEN
    RETURN;
END_IF
IF stLink.RxFill > MessageLen THEN
    MEMMOVE(destAddr := ADR(stLink.RxBuffer[0]),
            srcAddr  := ADR(stLink.RxBuffer[MessageLen]),
            n        := stLink.RxFill - MessageLen);
END_IF
stLink.RxFill    := stLink.RxFill - MessageLen;
MessageLen       := 0;
MessageAvailable := FALSE;
Consume := TRUE;
END_METHOD

END_FUNCTION_BLOCK

// ---- Library/POU/VC_DecodeHeader.TcPOU
FUNCTION VC_DecodeHeader : ST_VC_Header
VAR_IN_OUT
    Buf   : ARRAY[*] OF BYTE;
END_VAR
VAR
    stHdr : ST_VC_Header;
    nPos  : UDINT;
END_VAR

nPos := 0;
VC_GetRaw(Buf := Buf, Pos := nPos, pDst := ADR(stHdr), Size := VC_HEADER_LEN);
VC_DecodeHeader := stHdr;

END_FUNCTION

// ---- Library/POU/VC_GetRaw.TcPOU
FUNCTION VC_GetRaw : BOOL
// Copies Size bytes from Buf[Pos..] to pDst and advances Pos. Bounds-checked.
VAR_IN_OUT
    Buf  : ARRAY[*] OF BYTE;
    Pos  : UDINT;
END_VAR
VAR_INPUT
    pDst : PVOID;
    Size : UDINT;
END_VAR
VAR
    nHigh : DINT;
END_VAR

IF Size = 0 THEN
    VC_GetRaw := TRUE;
    RETURN;
END_IF
nHigh := UPPER_BOUND(Buf, 1);
IF (LOWER_BOUND(Buf, 1) <> 0) OR (pDst = 0) OR (nHigh < 0) OR ((Pos + Size) > (DINT_TO_UDINT(nHigh) + 1)) THEN
    VC_GetRaw := FALSE;
    RETURN;
END_IF
MEMCPY(destAddr := pDst, srcAddr := ADR(Buf[Pos]), n := Size);
Pos := Pos + Size;
VC_GetRaw := TRUE;

END_FUNCTION

// ---- Library/POU/VC_PutString.TcPOU
FUNCTION VC_PutString : BOOL
// Writes a fixed-length wire string: Len bytes ASCII, padded with 0.
VAR_IN_OUT
    Buf   : ARRAY[*] OF BYTE;
    Pos   : UDINT;
END_VAR
VAR_IN_OUT CONSTANT
    Value : STRING;
END_VAR
VAR_INPUT
    Len   : UDINT;      // wire length N from the interface definition
END_VAR
VAR
    nHigh : DINT;
    nCopy : UDINT;
END_VAR

IF Len = 0 THEN
    VC_PutString := TRUE;
    RETURN;
END_IF
nHigh := UPPER_BOUND(Buf, 1);
IF (LOWER_BOUND(Buf, 1) <> 0) OR (nHigh < 0) OR ((Pos + Len) > (DINT_TO_UDINT(nHigh) + 1)) THEN
    VC_PutString := FALSE;
    RETURN;
END_IF
MEMSET(destAddr := ADR(Buf[Pos]), fillByte := 0, n := Len);
nCopy := MIN(INT_TO_UDINT(LEN(Value)), Len);
IF nCopy > 0 THEN
    MEMCPY(destAddr := ADR(Buf[Pos]), srcAddr := ADR(Value), n := nCopy);
END_IF
Pos := Pos + Len;
VC_PutString := TRUE;

END_FUNCTION

// ---- Library/POU/VC_PutUInt16.TcPOU
FUNCTION VC_PutUInt16 : BOOL
// Writes UInt16 (2 byte, little-endian) at Buf[Pos] and advances Pos.
VAR_IN_OUT
    Buf   : ARRAY[*] OF BYTE;
    Pos   : UDINT;
END_VAR
VAR_INPUT
    Value : UINT;
END_VAR

VC_PutUInt16 := VC_PutRaw(Buf := Buf, Pos := Pos, pSrc := ADR(Value), Size := 2);

END_FUNCTION

// ---- Library/POU/VC_PutRaw.TcPOU
FUNCTION VC_PutRaw : BOOL
// Copies Size bytes from pSrc into Buf[Pos..] and advances Pos. Bounds-checked.
VAR_IN_OUT
    Buf  : ARRAY[*] OF BYTE;
    Pos  : UDINT;
END_VAR
VAR_INPUT
    pSrc : PVOID;
    Size : UDINT;
END_VAR
VAR
    nHigh : DINT;
END_VAR

IF Size = 0 THEN
    VC_PutRaw := TRUE;
    RETURN;
END_IF
nHigh := UPPER_BOUND(Buf, 1);
IF (LOWER_BOUND(Buf, 1) <> 0) OR (pSrc = 0) OR (nHigh < 0) OR ((Pos + Size) > (DINT_TO_UDINT(nHigh) + 1)) THEN
    VC_PutRaw := FALSE;
    RETURN;
END_IF
MEMCPY(destAddr := ADR(Buf[Pos]), srcAddr := pSrc, n := Size);
Pos := Pos + Size;
VC_PutRaw := TRUE;

END_FUNCTION

// ---- Library/POU/VC_PutUInt32.TcPOU
FUNCTION VC_PutUInt32 : BOOL
// Writes UInt32 (4 byte, little-endian) at Buf[Pos] and advances Pos.
VAR_IN_OUT
    Buf   : ARRAY[*] OF BYTE;
    Pos   : UDINT;
END_VAR
VAR_INPUT
    Value : UDINT;
END_VAR

VC_PutUInt32 := VC_PutRaw(Buf := Buf, Pos := Pos, pSrc := ADR(Value), Size := 4);

END_FUNCTION

// ---- Library/POU/VC_MethodIndex.TcPOU
FUNCTION VC_MethodIndex : INT
// Returns the method index for MethodId/Provider, or -1.
VAR_INPUT
    MethodId : UINT;
    Provider : USINT;
END_VAR
VAR
    i : UINT;
END_VAR

VC_MethodIndex := -1;
i := 0;
WHILE (i < VC_METHOD_COUNT) AND (i < VC_MAX_METHODS) DO
    IF (VC_METHODS[i].MethodId = MethodId) AND (VC_METHODS[i].Provider = Provider) THEN
        VC_MethodIndex := UINT_TO_INT(i);
        RETURN;
    END_IF
    i := i + 1;
END_WHILE

END_FUNCTION

// ---- Library/POU/VC_EncodeHeader.TcPOU
FUNCTION VC_EncodeHeader : BOOL
// Beckhoff: little-endian, packed struct copied 1:1 (Bausteindesign section 11)
VAR_IN_OUT
    Buf  : ARRAY[*] OF BYTE;
END_VAR
VAR_INPUT
    Hdr  : ST_VC_Header;
END_VAR
VAR
    nPos : UDINT;
END_VAR

nPos := 0;
VC_EncodeHeader := VC_PutRaw(Buf := Buf, Pos := nPos, pSrc := ADR(Hdr), Size := VC_HEADER_LEN);

END_FUNCTION

// ---- Generated/POU_Generated/VC_Call_StartInspection.TcPOU
FUNCTION_BLOCK VC_Call_StartInspection
// GENERATED (vcgen template, Bausteindesign 10.1). Calls App method 10 StartInspection.
// PLCopen behaviour: rising edge Execute starts; Done/Error held while Execute, at least 1 cycle.
VAR_INPUT
    Execute   : BOOL;
    Abort     : BOOL;
    RecipeId  : UINT;
    PartId    : STRING(31);
    TimeoutMs : UDINT;            // 0 = value from method table
END_VAR
VAR_IN_OUT
    Link      : ST_VC_LinkData;
END_VAR
VAR_OUTPUT
    Busy      : BOOL;
    Done      : BOOL;
    Error     : BOOL;
    ErrorId   : UINT;
    Result    : ST_VC_InspectionResult;
END_VAR
VAR CONSTANT
    METHOD_INDEX : UINT := VC_IDX_START_INSPECTION;
END_VAR
VAR
    rExec : R_TRIG;
    slot  : INT := -1;
    step  : INT;
    shown : BOOL;
    pos   : UDINT;
END_VAR

rExec(CLK := Execute);

CASE step OF
0:  // ready
    IF rExec.Q THEN
        Done := FALSE; Error := FALSE; ErrorId := 0;
        ErrorId := VC_IsCallable(Link := Link, MethodIndex := METHOD_INDEX);   // 0 = callable
        IF ErrorId = 0 THEN
            slot := VC_ReserveOutSlot(Link := Link, MethodIndex := METHOD_INDEX);
            IF slot < 0 THEN
                ErrorId := VC_STATUS_BUSY;
            END_IF
        END_IF
        IF ErrorId <> 0 THEN
            Error := TRUE; shown := FALSE; step := 2;
        ELSE
            // encode arguments (generated)
            pos := 0;
            VC_PutUInt16(Buf := Link.OutSlots[slot].Payload, Pos := pos, Value := RecipeId);
            VC_PutString(Buf := Link.OutSlots[slot].Payload, Pos := pos, Value := PartId, Len := 32);
            VC_SubmitOutSlot(Link := Link, Slot := slot, Len := pos, TimeoutMs := TimeoutMs);
            Busy := TRUE;
            step := 1;
        END_IF
    END_IF

1:  // call running
    IF (slot < 0) OR (Link.OutSlots[slot].State = VC_SS_FREE) THEN
        // slot lost (block was not called for > VC_OWNER_TIMEOUT_MS)
        Error := TRUE; ErrorId := VC_STATUS_INTERNAL_ERROR;
        slot := -1; Busy := FALSE; shown := FALSE;
        step := 2;
    ELSE
        Link.OutSlots[slot].OwnerSeenMs := Link.NowMs;
        IF Abort THEN
            VC_CancelOutSlot(Link := Link, Slot := slot);
        END_IF
        IF Link.OutSlots[slot].State = VC_SS_DONE THEN
            IF Link.OutSlots[slot].Status = VC_STATUS_OK THEN
                // decode result (generated)
                pos := 0;
                Result.Pass          := VC_GetBool(Buf := Link.OutSlots[slot].Payload, Pos := pos);
                Result.ErrorCode     := VC_GetInt32(Buf := Link.OutSlots[slot].Payload, Pos := pos);
                Result.MeasuredCount := VC_GetUInt16(Buf := Link.OutSlots[slot].Payload, Pos := pos);
                VC_GetFloat32Array(Buf := Link.OutSlots[slot].Payload, Pos := pos, Arr := Result.Measured, Count := 16);
                Done := TRUE;
            ELSE
                Error := TRUE;
                ErrorId := Link.OutSlots[slot].Status;
            END_IF
            VC_ReleaseOutSlot(Link := Link, Slot := slot);
            slot := -1; Busy := FALSE; shown := FALSE;
            step := 2;
        END_IF
    END_IF

2:  // show result, at least one cycle
    IF NOT Execute AND shown THEN
        Done := FALSE; Error := FALSE; ErrorId := 0;
        step := 0;
    END_IF
    shown := TRUE;
END_CASE

END_FUNCTION_BLOCK

// ---- Library/POU/VC_IsCallable.TcPOU
FUNCTION VC_IsCallable : UINT
// 0 = callable App method. Else 1 UnknownMethod, 8 ConnectionLost, 2 MethodIncompatible, 3 NotAllowed.
VAR_IN_OUT
    Link        : ST_VC_LinkData;
END_VAR
VAR_INPUT
    MethodIndex : UINT;
END_VAR

IF (MethodIndex >= VC_METHOD_COUNT) OR (MethodIndex >= VC_MAX_METHODS) THEN
    VC_IsCallable := VC_STATUS_UNKNOWN_METHOD;
ELSIF VC_METHODS[MethodIndex].Provider <> VC_PROVIDER_APP THEN
    VC_IsCallable := VC_STATUS_UNKNOWN_METHOD;
ELSIF NOT Link.Online THEN
    VC_IsCallable := VC_STATUS_CONNECTION_LOST;
ELSIF Link.MethodState[MethodIndex] = 1 THEN
    VC_IsCallable := VC_STATUS_OK;
ELSIF Link.MethodState[MethodIndex] = 3 THEN
    VC_IsCallable := VC_STATUS_NOT_ALLOWED;
ELSE
    VC_IsCallable := VC_STATUS_METHOD_INCOMPATIBLE;   // 0 unknown or 2 hash mismatch
END_IF

END_FUNCTION

// ---- Library/POU/VC_ReserveOutSlot.TcPOU
FUNCTION VC_ReserveOutSlot : INT
// First FREE out slot -> RESERVED. Returns slot or -1.
VAR_IN_OUT
    Link        : ST_VC_LinkData;
END_VAR
VAR_INPUT
    MethodIndex : UINT;
END_VAR
VAR
    i : UINT;
END_VAR

VC_ReserveOutSlot := -1;
FOR i := 0 TO VC_MAX_CALLS - 1 DO
    IF Link.OutSlots[i].State = VC_SS_FREE THEN
        Link.OutSlots[i].State       := VC_SS_RESERVED;
        Link.OutSlots[i].MethodIndex := MethodIndex;
        Link.OutSlots[i].OwnerSeenMs := Link.NowMs;
        Link.OutSlots[i].CallId      := 0;
        Link.OutSlots[i].Status      := VC_STATUS_OK;
        Link.OutSlots[i].PayloadLen  := 0;
        VC_ReserveOutSlot := UINT_TO_INT(i);
        RETURN;
    END_IF
END_FOR

END_FUNCTION

// ---- Library/POU/VC_SubmitOutSlot.TcPOU
FUNCTION VC_SubmitOutSlot : BOOL
// RESERVED -> TX_PENDING. Assigns CallId. TimeoutMs = 0 takes the table value.
VAR_IN_OUT
    Link      : ST_VC_LinkData;
END_VAR
VAR_INPUT
    Slot      : INT;
    Len       : UDINT;
    TimeoutMs : UDINT;
END_VAR
VAR
    nIdx : UINT;
END_VAR

VC_SubmitOutSlot := FALSE;
IF (Slot < 0) OR (Slot >= UINT_TO_INT(VC_MAX_CALLS)) THEN
    RETURN;
END_IF
IF Link.OutSlots[Slot].State <> VC_SS_RESERVED THEN
    RETURN;
END_IF
nIdx := Link.OutSlots[Slot].MethodIndex;

// Guard against generator / table mismatch
IF Len <> VC_METHODS[nIdx].ArgsLen THEN
    Link.OutSlots[Slot].Status     := VC_STATUS_INVALID_PAYLOAD;
    Link.OutSlots[Slot].PayloadLen := 0;
    Link.OutSlots[Slot].State      := VC_SS_DONE;
    RETURN;
END_IF

IF (Link.NextCallId = 0) OR (Link.NextCallId > 16#7FFFFFFF) THEN
    Link.NextCallId := 1;
END_IF
Link.OutSlots[Slot].CallId := Link.NextCallId;
Link.NextCallId := Link.NextCallId + 1;
IF Link.NextCallId > 16#7FFFFFFF THEN
    Link.NextCallId := 1;
END_IF

Link.OutSlots[Slot].PayloadLen := Len;
IF TimeoutMs = 0 THEN
    Link.OutSlots[Slot].TimeoutMs := VC_METHODS[nIdx].TimeoutMs;
ELSE
    Link.OutSlots[Slot].TimeoutMs := TimeoutMs;
END_IF
Link.OutSlots[Slot].StartMs := Link.NowMs;
Link.OutSlots[Slot].State   := VC_SS_TX_PENDING;
VC_SubmitOutSlot := TRUE;

END_FUNCTION

// ---- Library/POU/VC_CancelOutSlot.TcPOU
FUNCTION VC_CancelOutSlot : BOOL
// RESERVED/TX_PENDING -> DONE (Cancelled); SENT -> CANCEL_PENDING (Cancelled)
VAR_IN_OUT
    Link : ST_VC_LinkData;
END_VAR
VAR_INPUT
    Slot : INT;
END_VAR

VC_CancelOutSlot := FALSE;
IF (Slot < 0) OR (Slot >= UINT_TO_INT(VC_MAX_CALLS)) THEN
    RETURN;
END_IF
CASE Link.OutSlots[Slot].State OF
    VC_SS_RESERVED, VC_SS_TX_PENDING:
        Link.OutSlots[Slot].Status     := VC_STATUS_CANCELLED;
        Link.OutSlots[Slot].PayloadLen := 0;
        Link.OutSlots[Slot].State      := VC_SS_DONE;
        VC_CancelOutSlot := TRUE;
    VC_SS_SENT:
        Link.OutSlots[Slot].Status     := VC_STATUS_CANCELLED;
        Link.OutSlots[Slot].PayloadLen := 0;
        Link.OutSlots[Slot].State      := VC_SS_CANCEL_PENDING;
        VC_CancelOutSlot := TRUE;
END_CASE

END_FUNCTION

// ---- Library/POU/VC_GetBool.TcPOU
FUNCTION VC_GetBool : BOOL
// Reads Bool (1 byte, little-endian) from Buf[Pos] and advances Pos.
VAR_IN_OUT
    Buf   : ARRAY[*] OF BYTE;
    Pos   : UDINT;
END_VAR
VAR
    nByte : BYTE;
END_VAR

nByte := 0;
VC_GetRaw(Buf := Buf, Pos := Pos, pDst := ADR(nByte), Size := 1);
VC_GetBool := (nByte <> 0);

END_FUNCTION

// ---- Library/POU/VC_GetInt32.TcPOU
FUNCTION VC_GetInt32 : DINT
// Reads Int32 (4 byte, little-endian) from Buf[Pos] and advances Pos.
VAR_IN_OUT
    Buf   : ARRAY[*] OF BYTE;
    Pos   : UDINT;
END_VAR
VAR
    nVal : DINT;
END_VAR

nVal := 0;
VC_GetRaw(Buf := Buf, Pos := Pos, pDst := ADR(nVal), Size := 4);
VC_GetInt32 := nVal;

END_FUNCTION

// ---- Library/POU/VC_GetUInt16.TcPOU
FUNCTION VC_GetUInt16 : UINT
// Reads UInt16 (2 byte, little-endian) from Buf[Pos] and advances Pos.
VAR_IN_OUT
    Buf   : ARRAY[*] OF BYTE;
    Pos   : UDINT;
END_VAR
VAR
    nVal : UINT;
END_VAR

nVal := 0;
VC_GetRaw(Buf := Buf, Pos := Pos, pDst := ADR(nVal), Size := 2);
VC_GetUInt16 := nVal;

END_FUNCTION

// ---- Library/POU/VC_GetFloat32Array.TcPOU
FUNCTION VC_GetFloat32Array : BOOL
VAR_IN_OUT
    Buf   : ARRAY[*] OF BYTE;
    Pos   : UDINT;
    Arr   : ARRAY[*] OF REAL;
END_VAR
VAR_INPUT
    Count : UDINT;
END_VAR
VAR
    nLow  : DINT;
END_VAR

nLow := LOWER_BOUND(Arr, 1);
IF (UPPER_BOUND(Arr, 1) - nLow + 1) < UDINT_TO_DINT(Count) THEN
    VC_GetFloat32Array := FALSE;
    RETURN;
END_IF
VC_GetFloat32Array := VC_GetRaw(Buf := Buf, Pos := Pos, pDst := ADR(Arr[nLow]), Size := Count * 4);

END_FUNCTION

// ---- Library/POU/VC_ReleaseOutSlot.TcPOU
FUNCTION VC_ReleaseOutSlot : BOOL
VAR_IN_OUT
    Link : ST_VC_LinkData;
END_VAR
VAR_INPUT
    Slot : INT;
END_VAR

VC_ReleaseOutSlot := FALSE;
IF (Slot < 0) OR (Slot >= UINT_TO_INT(VC_MAX_CALLS)) THEN
    RETURN;
END_IF
Link.OutSlots[Slot].State      := VC_SS_FREE;
Link.OutSlots[Slot].Status     := VC_STATUS_OK;
Link.OutSlots[Slot].PayloadLen := 0;
VC_ReleaseOutSlot := TRUE;

END_FUNCTION

// ---- Generated/POU_Generated/VC_Handle_MoveToPosition.TcPOU
FUNCTION_BLOCK VC_Handle_MoveToPosition
// GENERATED (vcgen template, Bausteindesign 10.2). Provides PLC method 600 MoveToPosition.
// Call every cycle. NewRequest stays TRUE until a rising edge of Respond.
VAR_INPUT
    Respond        : BOOL;
    ResponseStatus : UINT;        // 0 or business error code (>= 5000 for project errors)
    Result         : ST_VC_MoveToPositionResult;
END_VAR
VAR_IN_OUT
    Link           : ST_VC_LinkData;
END_VAR
VAR_OUTPUT
    NewRequest      : BOOL;
    Args            : ST_VC_MoveToPositionArgs;
    CancelRequested : BOOL;
END_VAR
VAR CONSTANT
    METHOD_INDEX : UINT := VC_IDX_MOVE_TO_POSITION;
END_VAR
VAR
    rResp  : R_TRIG;
    slot   : INT := -1;
    callId : UDINT;
    pos    : UDINT;
END_VAR

Link.HandlerSeenMs[METHOD_INDEX] := Link.NowMs;   // handler is active
rResp(CLK := Respond);

IF slot < 0 THEN
    slot := VC_TakeInSlot(Link := Link, MethodIndex := METHOD_INDEX);   // REQUEST -> IN_PROGRESS
    IF slot >= 0 THEN
        callId := Link.InSlots[slot].CallId;
        pos := 0;
        Args.Position := VC_GetFloat64(Buf := Link.InSlots[slot].Payload, Pos := pos);   // generated
        NewRequest := TRUE;
    END_IF
END_IF

IF slot >= 0 THEN
    // slot lost (deadline, connection loss)?
    IF (Link.InSlots[slot].State <> VC_SS_IN_PROGRESS) OR (Link.InSlots[slot].CallId <> callId) THEN
        slot := -1; NewRequest := FALSE; CancelRequested := FALSE;
    ELSE
        CancelRequested := Link.InSlots[slot].CancelRequested;
        IF rResp.Q THEN
            pos := 0;
            IF ResponseStatus = VC_STATUS_OK THEN
                VC_PutBool(Buf := Link.InSlots[slot].Payload, Pos := pos, Value := Result.Accepted);   // generated
            END_IF
            VC_CompleteInSlot(Link := Link, Slot := slot, Status := ResponseStatus, Len := pos);   // -> RESPONSE_READY
            slot := -1; NewRequest := FALSE; CancelRequested := FALSE;
        END_IF
    END_IF
END_IF

END_FUNCTION_BLOCK

// ---- Library/POU/VC_TakeInSlot.TcPOU
FUNCTION VC_TakeInSlot : INT
// Oldest REQUEST slot of this method -> IN_PROGRESS. Returns slot or -1.
VAR_IN_OUT
    Link        : ST_VC_LinkData;
END_VAR
VAR_INPUT
    MethodIndex : UINT;
END_VAR
VAR
    i       : UINT;
    nBest   : INT;
    nAge    : UDINT;
    nBestAge: UDINT;
END_VAR

nBest := -1;
nBestAge := 0;
FOR i := 0 TO VC_MAX_CALLS - 1 DO
    IF (Link.InSlots[i].State = VC_SS_REQUEST) AND (Link.InSlots[i].MethodIndex = MethodIndex) THEN
        nAge := Link.NowMs - Link.InSlots[i].ReceivedMs;
        IF (nBest < 0) OR (nAge > nBestAge) THEN
            nBest := UINT_TO_INT(i);
            nBestAge := nAge;
        END_IF
    END_IF
END_FOR
IF nBest >= 0 THEN
    Link.InSlots[nBest].State := VC_SS_IN_PROGRESS;
END_IF
VC_TakeInSlot := nBest;

END_FUNCTION

// ---- Library/POU/VC_GetFloat64.TcPOU
FUNCTION VC_GetFloat64 : LREAL
// Reads Float64 (8 byte, little-endian) from Buf[Pos] and advances Pos.
VAR_IN_OUT
    Buf   : ARRAY[*] OF BYTE;
    Pos   : UDINT;
END_VAR
VAR
    nVal : LREAL;
END_VAR

nVal := 0;
VC_GetRaw(Buf := Buf, Pos := Pos, pDst := ADR(nVal), Size := 8);
VC_GetFloat64 := nVal;

END_FUNCTION

// ---- Library/POU/VC_PutBool.TcPOU
FUNCTION VC_PutBool : BOOL
// Writes Bool (1 byte, little-endian) at Buf[Pos] and advances Pos.
VAR_IN_OUT
    Buf   : ARRAY[*] OF BYTE;
    Pos   : UDINT;
END_VAR
VAR_INPUT
    Value : BOOL;
END_VAR
VAR
    nByte : BYTE;
END_VAR

nByte := BOOL_TO_BYTE(Value);   // wire: 0 or 1
VC_PutBool := VC_PutRaw(Buf := Buf, Pos := Pos, pSrc := ADR(nByte), Size := 1);

END_FUNCTION

// ---- Library/POU/VC_CompleteInSlot.TcPOU
FUNCTION VC_CompleteInSlot : BOOL
// IN_PROGRESS -> RESPONSE_READY. Len is ignored (0) when Status <> 0.
VAR_IN_OUT
    Link   : ST_VC_LinkData;
END_VAR
VAR_INPUT
    Slot   : INT;
    Status : UINT;
    Len    : UDINT;
END_VAR
VAR
    nIdx    : UINT;
    nStatus : UINT;
END_VAR

VC_CompleteInSlot := FALSE;
IF (Slot < 0) OR (Slot >= UINT_TO_INT(VC_MAX_CALLS)) THEN
    RETURN;
END_IF
IF Link.InSlots[Slot].State <> VC_SS_IN_PROGRESS THEN
    RETURN;
END_IF
nIdx := Link.InSlots[Slot].MethodIndex;
nStatus := Status;
IF (nStatus = VC_STATUS_OK) AND (Len <> VC_METHODS[nIdx].ResultLen) THEN
    nStatus := VC_STATUS_INTERNAL_ERROR;     // generator / table mismatch
END_IF
Link.InSlots[Slot].Status := nStatus;
IF nStatus = VC_STATUS_OK THEN
    Link.InSlots[Slot].PayloadLen := Len;
ELSE
    Link.InSlots[Slot].PayloadLen := 0;
END_IF
Link.InSlots[Slot].State := VC_SS_RESPONSE_READY;
VC_CompleteInSlot := TRUE;

END_FUNCTION

// ---- Generated/POU_Generated/VC_Handle_ReportModuleState.TcPOU
FUNCTION_BLOCK VC_Handle_ReportModuleState
// GENERATED (vcgen template). Provides PLC method 500 ReportModuleState (no result payload).
VAR_INPUT
    Respond        : BOOL;
    ResponseStatus : UINT;
END_VAR
VAR_IN_OUT
    Link           : ST_VC_LinkData;
END_VAR
VAR_OUTPUT
    NewRequest      : BOOL;
    Args            : ST_VC_ReportModuleStateArgs;
    CancelRequested : BOOL;
END_VAR
VAR CONSTANT
    METHOD_INDEX : UINT := VC_IDX_REPORT_MODULE_STATE;
END_VAR
VAR
    rResp  : R_TRIG;
    slot   : INT := -1;
    callId : UDINT;
    pos    : UDINT;
END_VAR

Link.HandlerSeenMs[METHOD_INDEX] := Link.NowMs;
rResp(CLK := Respond);

IF slot < 0 THEN
    slot := VC_TakeInSlot(Link := Link, MethodIndex := METHOD_INDEX);
    IF slot >= 0 THEN
        callId := Link.InSlots[slot].CallId;
        pos := 0;
        Args.State   := VC_GetUInt16(Buf := Link.InSlots[slot].Payload, Pos := pos);
        Args.AlarmId := VC_GetInt32(Buf := Link.InSlots[slot].Payload, Pos := pos);
        NewRequest := TRUE;
    END_IF
END_IF

IF slot >= 0 THEN
    IF (Link.InSlots[slot].State <> VC_SS_IN_PROGRESS) OR (Link.InSlots[slot].CallId <> callId) THEN
        slot := -1; NewRequest := FALSE; CancelRequested := FALSE;
    ELSE
        CancelRequested := Link.InSlots[slot].CancelRequested;
        IF rResp.Q THEN
            VC_CompleteInSlot(Link := Link, Slot := slot, Status := ResponseStatus, Len := 0);
            slot := -1; NewRequest := FALSE; CancelRequested := FALSE;
        END_IF
    END_IF
END_IF

END_FUNCTION_BLOCK

// ---- Library/POU/VC_GetFloat32.TcPOU
FUNCTION VC_GetFloat32 : REAL
// Reads Float32 (4 byte, little-endian) from Buf[Pos] and advances Pos.
VAR_IN_OUT
    Buf   : ARRAY[*] OF BYTE;
    Pos   : UDINT;
END_VAR
VAR
    nVal : REAL;
END_VAR

nVal := 0;
VC_GetRaw(Buf := Buf, Pos := Pos, pDst := ADR(nVal), Size := 4);
VC_GetFloat32 := nVal;

END_FUNCTION

// ---- Library/POU/VC_GetInt16.TcPOU
FUNCTION VC_GetInt16 : INT
// Reads Int16 (2 byte, little-endian) from Buf[Pos] and advances Pos.
VAR_IN_OUT
    Buf   : ARRAY[*] OF BYTE;
    Pos   : UDINT;
END_VAR
VAR
    nVal : INT;
END_VAR

nVal := 0;
VC_GetRaw(Buf := Buf, Pos := Pos, pDst := ADR(nVal), Size := 2);
VC_GetInt16 := nVal;

END_FUNCTION

// ---- Library/POU/VC_GetInt64.TcPOU
FUNCTION VC_GetInt64 : LINT
// Reads Int64 (8 byte, little-endian) from Buf[Pos] and advances Pos.
VAR_IN_OUT
    Buf   : ARRAY[*] OF BYTE;
    Pos   : UDINT;
END_VAR
VAR
    nVal : LINT;
END_VAR

nVal := 0;
VC_GetRaw(Buf := Buf, Pos := Pos, pDst := ADR(nVal), Size := 8);
VC_GetInt64 := nVal;

END_FUNCTION

// ---- Library/POU/VC_GetInt8.TcPOU
FUNCTION VC_GetInt8 : SINT
// Reads Int8 (1 byte, little-endian) from Buf[Pos] and advances Pos.
VAR_IN_OUT
    Buf   : ARRAY[*] OF BYTE;
    Pos   : UDINT;
END_VAR
VAR
    nVal : SINT;
END_VAR

nVal := 0;
VC_GetRaw(Buf := Buf, Pos := Pos, pDst := ADR(nVal), Size := 1);
VC_GetInt8 := nVal;

END_FUNCTION

// ---- Library/POU/VC_GetString.TcPOU
FUNCTION VC_GetString : STRING(255)
// Reads a fixed-length wire string of Len bytes. Assign the result to STRING(Len-1).
VAR_IN_OUT
    Buf   : ARRAY[*] OF BYTE;
    Pos   : UDINT;
END_VAR
VAR_INPUT
    Len   : UDINT;
END_VAR
VAR
    sTmp  : STRING(255);
    nHigh : DINT;
END_VAR

MEMSET(destAddr := ADR(sTmp), fillByte := 0, n := SIZEOF(sTmp));
nHigh := UPPER_BOUND(Buf, 1);
IF (Len > 0) AND (LOWER_BOUND(Buf, 1) = 0) AND (nHigh >= 0) AND ((Pos + Len) <= (DINT_TO_UDINT(nHigh) + 1)) THEN
    MEMCPY(destAddr := ADR(sTmp), srcAddr := ADR(Buf[Pos]), n := MIN(Len, 255));
    Pos := Pos + Len;
END_IF
VC_GetString := sTmp;

END_FUNCTION

// ---- Library/POU/VC_GetUInt32.TcPOU
FUNCTION VC_GetUInt32 : UDINT
// Reads UInt32 (4 byte, little-endian) from Buf[Pos] and advances Pos.
VAR_IN_OUT
    Buf   : ARRAY[*] OF BYTE;
    Pos   : UDINT;
END_VAR
VAR
    nVal : UDINT;
END_VAR

nVal := 0;
VC_GetRaw(Buf := Buf, Pos := Pos, pDst := ADR(nVal), Size := 4);
VC_GetUInt32 := nVal;

END_FUNCTION

// ---- Library/POU/VC_GetUInt64.TcPOU
FUNCTION VC_GetUInt64 : ULINT
// Reads UInt64 (8 byte, little-endian) from Buf[Pos] and advances Pos.
VAR_IN_OUT
    Buf   : ARRAY[*] OF BYTE;
    Pos   : UDINT;
END_VAR
VAR
    nVal : ULINT;
END_VAR

nVal := 0;
VC_GetRaw(Buf := Buf, Pos := Pos, pDst := ADR(nVal), Size := 8);
VC_GetUInt64 := nVal;

END_FUNCTION

// ---- Library/POU/VC_GetUInt8.TcPOU
FUNCTION VC_GetUInt8 : USINT
// Reads UInt8 (1 byte, little-endian) from Buf[Pos] and advances Pos.
VAR_IN_OUT
    Buf   : ARRAY[*] OF BYTE;
    Pos   : UDINT;
END_VAR
VAR
    nVal : USINT;
END_VAR

nVal := 0;
VC_GetRaw(Buf := Buf, Pos := Pos, pDst := ADR(nVal), Size := 1);
VC_GetUInt8 := nVal;

END_FUNCTION

// ---- Library/POU/VC_PutFloat32.TcPOU
FUNCTION VC_PutFloat32 : BOOL
// Writes Float32 (4 byte, little-endian) at Buf[Pos] and advances Pos.
VAR_IN_OUT
    Buf   : ARRAY[*] OF BYTE;
    Pos   : UDINT;
END_VAR
VAR_INPUT
    Value : REAL;
END_VAR

VC_PutFloat32 := VC_PutRaw(Buf := Buf, Pos := Pos, pSrc := ADR(Value), Size := 4);

END_FUNCTION

// ---- Library/POU/VC_PutFloat32Array.TcPOU
FUNCTION VC_PutFloat32Array : BOOL
VAR_IN_OUT
    Buf   : ARRAY[*] OF BYTE;
    Pos   : UDINT;
    Arr   : ARRAY[*] OF REAL;
END_VAR
VAR_INPUT
    Count : UDINT;
END_VAR
VAR
    nLow  : DINT;
END_VAR

nLow := LOWER_BOUND(Arr, 1);
IF (UPPER_BOUND(Arr, 1) - nLow + 1) < UDINT_TO_DINT(Count) THEN
    VC_PutFloat32Array := FALSE;
    RETURN;
END_IF
VC_PutFloat32Array := VC_PutRaw(Buf := Buf, Pos := Pos, pSrc := ADR(Arr[nLow]), Size := Count * 4);

END_FUNCTION

// ---- Library/POU/VC_PutFloat64.TcPOU
FUNCTION VC_PutFloat64 : BOOL
// Writes Float64 (8 byte, little-endian) at Buf[Pos] and advances Pos.
VAR_IN_OUT
    Buf   : ARRAY[*] OF BYTE;
    Pos   : UDINT;
END_VAR
VAR_INPUT
    Value : LREAL;
END_VAR

VC_PutFloat64 := VC_PutRaw(Buf := Buf, Pos := Pos, pSrc := ADR(Value), Size := 8);

END_FUNCTION

// ---- Library/POU/VC_PutInt16.TcPOU
FUNCTION VC_PutInt16 : BOOL
// Writes Int16 (2 byte, little-endian) at Buf[Pos] and advances Pos.
VAR_IN_OUT
    Buf   : ARRAY[*] OF BYTE;
    Pos   : UDINT;
END_VAR
VAR_INPUT
    Value : INT;
END_VAR

VC_PutInt16 := VC_PutRaw(Buf := Buf, Pos := Pos, pSrc := ADR(Value), Size := 2);

END_FUNCTION

// ---- Library/POU/VC_PutInt32.TcPOU
FUNCTION VC_PutInt32 : BOOL
// Writes Int32 (4 byte, little-endian) at Buf[Pos] and advances Pos.
VAR_IN_OUT
    Buf   : ARRAY[*] OF BYTE;
    Pos   : UDINT;
END_VAR
VAR_INPUT
    Value : DINT;
END_VAR

VC_PutInt32 := VC_PutRaw(Buf := Buf, Pos := Pos, pSrc := ADR(Value), Size := 4);

END_FUNCTION

// ---- Library/POU/VC_PutInt64.TcPOU
FUNCTION VC_PutInt64 : BOOL
// Writes Int64 (8 byte, little-endian) at Buf[Pos] and advances Pos.
VAR_IN_OUT
    Buf   : ARRAY[*] OF BYTE;
    Pos   : UDINT;
END_VAR
VAR_INPUT
    Value : LINT;
END_VAR

VC_PutInt64 := VC_PutRaw(Buf := Buf, Pos := Pos, pSrc := ADR(Value), Size := 8);

END_FUNCTION

// ---- Library/POU/VC_PutInt8.TcPOU
FUNCTION VC_PutInt8 : BOOL
// Writes Int8 (1 byte, little-endian) at Buf[Pos] and advances Pos.
VAR_IN_OUT
    Buf   : ARRAY[*] OF BYTE;
    Pos   : UDINT;
END_VAR
VAR_INPUT
    Value : SINT;
END_VAR

VC_PutInt8 := VC_PutRaw(Buf := Buf, Pos := Pos, pSrc := ADR(Value), Size := 1);

END_FUNCTION

// ---- Library/POU/VC_PutUInt64.TcPOU
FUNCTION VC_PutUInt64 : BOOL
// Writes UInt64 (8 byte, little-endian) at Buf[Pos] and advances Pos.
VAR_IN_OUT
    Buf   : ARRAY[*] OF BYTE;
    Pos   : UDINT;
END_VAR
VAR_INPUT
    Value : ULINT;
END_VAR

VC_PutUInt64 := VC_PutRaw(Buf := Buf, Pos := Pos, pSrc := ADR(Value), Size := 8);

END_FUNCTION

// ---- Library/POU/VC_PutUInt8.TcPOU
FUNCTION VC_PutUInt8 : BOOL
// Writes UInt8 (1 byte, little-endian) at Buf[Pos] and advances Pos.
VAR_IN_OUT
    Buf   : ARRAY[*] OF BYTE;
    Pos   : UDINT;
END_VAR
VAR_INPUT
    Value : USINT;
END_VAR

VC_PutUInt8 := VC_PutRaw(Buf := Buf, Pos := Pos, pSrc := ADR(Value), Size := 1);

END_FUNCTION

// ---- POUs/MAIN.TcPOU
PROGRAM MAIN
VAR
	btn:BOOL;
END_VAR


// 
// IF not btn THEN
// ADSLOGSTR( msgCtrlMask := ADSLOG_MSGTYPE_ERROR OR ADSLOG_MSGTYPE_LOG ,
//            msgFmtStr  := 'Hello %s',
//            strArg     := 'world!' );
// 		   btn :=TRUE;
// END_IF

END_PROGRAM

// ---- Test/POU/FB_VC_LinkTest.TcPOU
FUNCTION_BLOCK FB_VC_LinkTest
// Test harness: one link, one App call, two PLC handlers. Order per cycle: link first, then method blocks.
VAR_INPUT
    bEnable          : BOOL;
    nMode            : INT := 0;                    // 0 = PLC connects (VisionCore Listen), 1 = PLC listens
    sRemoteAddress   : STRING(15) := '127.0.0.1';   // VisionCore on the same PC
    nPort            : UINT := 5100;
    sClientId        : STRING(31) := 'Line1_Plc';   // must match VisionCore PlcLinkDevice config
    bStartInspection : BOOL;                        // set TRUE online -> one call
    bAbortInspection : BOOL;
    nRecipeId        : UINT := 1;
    sPartId          : STRING(31) := 'TEST_0001';
    bAcceptMove      : BOOL := TRUE;                // MoveToPosition answer
END_VAR
VAR_OUTPUT
    eLinkState     : E_VC_LinkState;
    bConnected     : BOOL;
    bOnline        : BOOL;
    bRestricted    : BOOL;
    nLinkErrorId   : UINT;
    bInspBusy      : BOOL;
    bInspDone      : BOOL;
    nInspErrorId   : UINT;
    stInspResult   : ST_VC_InspectionResult;
    nMoveRequests  : UDINT;
    lrLastPosition : LREAL;
    nStateReports  : UDINT;
    nVisionState   : UINT;
    nVisionAlarm   : DINT;
END_VAR
VAR
    fbLink        : VC_Link;
    fbInspect     : VC_Call_StartInspection;
    fbMove        : VC_Handle_MoveToPosition;
    fbModuleState : VC_Handle_ReportModuleState;
    bRespondMove  : BOOL;
    bRespondState : BOOL;
    stMoveResult  : ST_VC_MoveToPositionResult;
END_VAR

THIS^.RunLink();
THIS^.CallInspection();
THIS^.HandleMove();
THIS^.HandleModuleState();

METHOD PRIVATE CallInspection
fbInspect(Execute   := bStartInspection,
          Abort     := bAbortInspection,
          RecipeId  := nRecipeId,
          PartId    := sPartId,
          TimeoutMs := 0,
          Link      := GVL_VC.LinkData);
bInspBusy := fbInspect.Busy;
IF fbInspect.Busy THEN
    bInspDone    := FALSE;
    nInspErrorId := 0;
END_IF
IF fbInspect.Done THEN
    bInspDone        := TRUE;
    stInspResult     := fbInspect.Result;
    bStartInspection := FALSE;
ELSIF fbInspect.Error THEN
    nInspErrorId     := fbInspect.ErrorId;
    bStartInspection := FALSE;
END_IF
END_METHOD

METHOD PRIVATE HandleModuleState
fbModuleState(Respond        := bRespondState,
              ResponseStatus := VC_STATUS_OK,
              Link           := GVL_VC.LinkData);
IF fbModuleState.NewRequest AND NOT bRespondState THEN
    nVisionState  := fbModuleState.Args.State;     // -> PackML tags
    nVisionAlarm  := fbModuleState.Args.AlarmId;
    nStateReports := nStateReports + 1;
END_IF
bRespondState := fbModuleState.NewRequest AND NOT bRespondState;
END_METHOD

METHOD PRIVATE HandleMove
// Answers one cycle after NewRequest so Respond gets a clean rising edge.
stMoveResult.Accepted := bAcceptMove;
fbMove(Respond        := bRespondMove,
       ResponseStatus := SEL(fbMove.CancelRequested, VC_STATUS_OK, VC_STATUS_CANCELLED),
       Result         := stMoveResult,
       Link           := GVL_VC.LinkData);
IF fbMove.NewRequest AND NOT bRespondMove THEN
    lrLastPosition := fbMove.Args.Position;   // real cell: start axis here, answer when accepted
    nMoveRequests  := nMoveRequests + 1;
END_IF
bRespondMove := fbMove.NewRequest AND NOT bRespondMove;
END_METHOD

METHOD PRIVATE RunLink
fbLink(Enable        := bEnable,
       Mode          := nMode,
       RemoteAddress := sRemoteAddress,
       RemotePort    := nPort,
       LocalPort     := nPort,
       ClientId      := sClientId,
       Link          := GVL_VC.LinkData);
eLinkState   := fbLink.State;
bConnected   := fbLink.Connected;
bOnline      := fbLink.Online;
bRestricted  := fbLink.Restricted;
nLinkErrorId := fbLink.ErrorId;      // kept until ONLINE again
END_METHOD

END_FUNCTION_BLOCK

// ---- Test/POU/MAIN_1.TcPOU
PROGRAM MAIN_1
VAR
    fbCloseAll : FB_SocketCloseAll;   // closes stale sockets after download / restart
    bInitDone  : BOOL;
    bEnable    : BOOL := TRUE;
    fbTest     : FB_VC_LinkTest;
END_VAR

// Once at startup. NOTE: closes ALL TF6310 sockets of this runtime.
IF NOT bInitDone THEN
    fbCloseAll(sSrvNetId := '', bExecute := TRUE, tTimeout := T#5S);
    IF NOT fbCloseAll.bBusy THEN
        fbCloseAll(bExecute := FALSE);
        bInitDone := TRUE;
    END_IF
END_IF

fbTest(bEnable := bEnable AND bInitDone);

END_PROGRAM
